(* IEC 61131-3 sources: 2026_Projet_YGO_ExcavatriceDragage/ARCHIVES/Code/PLC_TESTS/CORE, 6 files *)

(* ---- FB_TranslationReportFinalizer.st ---- *)
// ═══════════════════════════════════════════════════════════════
// 🧪 FB_TranslationReportFinalizer — Rapport incrémental Translation
// ───────────────────────────────────────────────────────────────
// 🎯 Responsabilité UNIQUE : enregistrer les verdicts réels et finaliser
//    un rapport borné. Aucun parcours du graphe de transitions.
// ═══════════════════════════════════════════════════════════════

FUNCTION_BLOCK PUBLIC FB_TranslationReportFinalizer
VAR_INPUT
    RunStart        : BOOL;
    RequestedCaseId : INT;
    Busy            : BOOL;
    StepVerdict         : BOOL;
    StepId              : INT;
    StepCaseId          : INT;
    StepPassed          : BOOL;
    StepFailReason      : E_TestFailReason;
    StepFailedCheckIdx  : INT;
    StepDuration        : TIME;
    StepObservedBool    : BOOL;
    StepObservedDint    : DINT;
    StepObservedReal    : REAL;
    Finalize       : BOOL;
    TerminalState  : E_TestTerminalState;
    ErrorCode      : INT;
    ErrorMessage   : STRING(160);
END_VAR
VAR_IN_OUT
    StepTable : ARRAY[1..GVL_PLC_Tests_Const.MaxSteps]     OF ST_TestStepConfig;
    CaseTable : ARRAY[1..GVL_PLC_Tests_Const.MaxTestCases] OF ST_TestCaseConfig;
    Report    : ST_TestSuiteReport;
    Result    : ST_TranslationTestResult;
END_VAR
VAR
    Idx             : INT;
    CaseIdx         : INT;
    CasesTotalLocal : INT;
    CasesPassedLocal: INT;
    CasesFailedLocal: INT;
    FirstFailedCase : INT;
    ReasonText      : STRING(20);
    EntryText       : STRING(80);
END_VAR
// === IMPLEMENTATION ===
IF RunStart THEN
    Report.Name := 'Translation Validation';
    Report.InProgress := TRUE;
    Report.AllPassed := FALSE;
    Report.AnyFailed := FALSE;
    Report.Aborted := FALSE;
    Report.TerminalState := E_TestTerminalState.TEST_TERMINAL_NONE;
    Report.ErrorCode := 0;
    Report.ErrorMessage := '';
    Report.FailedTestCase := 0;
    Report.FailureSummary := '';
    Report.CurrentStepId := 0;
    Report.CurrentCaseId := 0;
    Report.Duration := T#0s;
    Report.RunCounter := Report.RunCounter + 1;
    FOR Idx := 1 TO GVL_PLC_Tests_Const.MaxSteps DO
        Report.Steps[Idx].Executed := FALSE;
        Report.Steps[Idx].Passed := FALSE;
        Report.Steps[Idx].FailReason := E_TestFailReason.FAIL_NONE;
        Report.Steps[Idx].FailedCheckIdx := 0;
        Report.Steps[Idx].FailedInvariantId := 0;
        Report.Steps[Idx].Duration := T#0s;
    END_FOR;
    FOR Idx := 1 TO GVL_PLC_Tests_Const.MaxTestCases DO
        Report.Cases[Idx].Name := CaseTable[Idx].Name;
        Report.Cases[Idx].Executed := FALSE;
        Report.Cases[Idx].Ok := FALSE;
        Report.Cases[Idx].FailedStepId := 0;
        Report.Cases[Idx].FailReason := E_TestFailReason.FAIL_NONE;
        Report.Cases[Idx].Duration := T#0s;
    END_FOR;
    Result.TerminalState := E_TestTerminalState.TEST_TERMINAL_NONE;
    Result.RequestedCaseId := RequestedCaseId;
    Result.ExecutedCaseId := 0;
    Result.AllPassed := FALSE;
    Result.AnyFailed := FALSE;
    Result.FailedCaseId := 0;
    Result.FailedCaseName := '';
    Result.FailReason := E_TestFailReason.FAIL_NONE;
    Result.ErrorCode := 0;
    Result.ErrorMessage := '';
    Result.CasesTotal := 0;
    Result.CasesPassed := 0;
    Result.CasesFailed := 0;
    Result.Duration := T#0s;
    Result.RunCounter := Report.RunCounter;
END_IF;

IF Busy THEN
    Report.Duration := Report.Duration + UDINT_TO_TIME(INT_TO_UDINT(GVL_PLC_Tests_Const.TaskCycleMs));
END_IF;

// 🧾 Agrégation incrémentale : validation séparée avant toute indexation.
IF StepVerdict THEN
    IF StepId < 1 OR StepId > GVL_PLC_Tests_Const.MaxSteps THEN
        Report.ErrorCode := 1050;
        Report.ErrorMessage := 'Verdict StepId hors limites';
        Report.AnyFailed := TRUE;
        RETURN;
    END_IF;
    Report.Steps[StepId].Executed := TRUE;
    Report.Steps[StepId].Passed := StepPassed;
    Report.Steps[StepId].FailReason := StepFailReason;
    Report.Steps[StepId].FailedCheckIdx := StepFailedCheckIdx;
    Report.Steps[StepId].Duration := StepDuration;
    Report.Steps[StepId].ObservedBool := StepObservedBool;
    Report.Steps[StepId].ObservedDint := StepObservedDint;
    Report.Steps[StepId].ObservedReal := StepObservedReal;
    Report.CurrentStepId := StepId;
    Report.CurrentCaseId := StepCaseId;

    IF StepCaseId >= 1 THEN
        IF StepCaseId <= GVL_PLC_Tests_Const.MaxTestCases THEN
        IF NOT Report.Cases[StepCaseId].Executed THEN
            Report.Cases[StepCaseId].Executed := TRUE;
            Report.Cases[StepCaseId].Ok := TRUE;
        END_IF;
        Report.Cases[StepCaseId].Duration := Report.Cases[StepCaseId].Duration + StepDuration;
        IF NOT StepPassed THEN
            Report.Cases[StepCaseId].Ok := FALSE;
            IF Report.Cases[StepCaseId].FailedStepId = 0 THEN
                Report.Cases[StepCaseId].FailedStepId := StepId;
                Report.Cases[StepCaseId].FailReason := StepFailReason;
            END_IF;
        END_IF;
        ELSE
            Report.ErrorCode := 1051;
            Report.ErrorMessage := 'Verdict CaseId hors limites';
            Report.AnyFailed := TRUE;
        END_IF;
    ELSE
        Report.ErrorCode := 1051;
        Report.ErrorMessage := 'Verdict CaseId hors limites';
        Report.AnyFailed := TRUE;
    END_IF;
END_IF;

IF Finalize THEN
    Report.InProgress := FALSE;
    Report.TerminalState := TerminalState;
    Report.ErrorCode := ErrorCode;
    Report.ErrorMessage := ErrorMessage;
    Report.Aborted := (TerminalState = E_TestTerminalState.TEST_TERMINAL_ABORTED);
    CasesTotalLocal := 0;
    CasesPassedLocal := 0;
    CasesFailedLocal := 0;
    FirstFailedCase := 0;
    Report.FailureSummary := '';

    FOR CaseIdx := 1 TO GVL_PLC_Tests_Const.MaxTestCases DO
        IF Report.Cases[CaseIdx].Executed THEN
            CasesTotalLocal := CasesTotalLocal + 1;
            IF Report.Cases[CaseIdx].Ok THEN
                CasesPassedLocal := CasesPassedLocal + 1;
            ELSE
                CasesFailedLocal := CasesFailedLocal + 1;
                IF FirstFailedCase = 0 THEN FirstFailedCase := CaseIdx; END_IF;
                CASE Report.Cases[CaseIdx].FailReason OF
                    E_TestFailReason.FAIL_TIMEOUT: ReasonText := 'FAIL_TIMEOUT';
                    E_TestFailReason.FAIL_CHECK: ReasonText := 'FAIL_CHECK';
                    E_TestFailReason.FAIL_INVARIANT: ReasonText := 'FAIL_INVARIANT';
                    E_TestFailReason.FAIL_WINDOW_EARLY: ReasonText := 'FAIL_WINDOW_EARLY';
                    E_TestFailReason.FAIL_ABORTED: ReasonText := 'FAIL_ABORTED';
                ELSE ReasonText := 'FAIL_NONE';
                END_CASE;
                EntryText := CONCAT(Report.Cases[CaseIdx].Name, ' (step ');
                EntryText := CONCAT(EntryText, INT_TO_STRING(Report.Cases[CaseIdx].FailedStepId));
                EntryText := CONCAT(EntryText, '): ');
                EntryText := CONCAT(EntryText, ReasonText);
                IF Report.FailureSummary = '' THEN
                    Report.FailureSummary := EntryText;
                ELSE
                    Report.FailureSummary := CONCAT(Report.FailureSummary, ' | ');
                    Report.FailureSummary := CONCAT(Report.FailureSummary, EntryText);
                END_IF;
            END_IF;
        END_IF;
    END_FOR;

    Report.AllPassed := (TerminalState = E_TestTerminalState.TEST_TERMINAL_DONE)
                     AND (CasesTotalLocal > 0)
                     AND (CasesFailedLocal = 0);
    Report.AnyFailed := NOT Report.AllPassed;
    Report.FailedTestCase := FirstFailedCase;

    Result.TerminalState := TerminalState;
    Result.RequestedCaseId := RequestedCaseId;
    Result.ExecutedCaseId := Report.CurrentCaseId;
    Result.AllPassed := Report.AllPassed;
    Result.AnyFailed := Report.AnyFailed;
    Result.FailedCaseId := FirstFailedCase;
    IF FirstFailedCase > 0 THEN
        Result.FailedCaseName := Report.Cases[FirstFailedCase].Name;
        Result.FailReason := Report.Cases[FirstFailedCase].FailReason;
    ELSE
        Result.FailedCaseName := '';
        Result.FailReason := E_TestFailReason.FAIL_NONE;
    END_IF;
    Result.ErrorCode := ErrorCode;
    Result.ErrorMessage := ErrorMessage;
    Result.CasesTotal := CasesTotalLocal;
    Result.CasesPassed := CasesPassedLocal;
    Result.CasesFailed := CasesFailedLocal;
    Result.Duration := Report.Duration;
    Result.RunCounter := Report.RunCounter;
END_IF;

(* ---- FB_TranslationStepExecutor.st ---- *)
// ═══════════════════════════════════════════════════════════════
// 🧪 FB_TranslationStepExecutor — Exécution étape/check Translation M3
// ───────────────────────────────────────────────────────────────
// 🎯 Responsabilité UNIQUE : faire progresser UNE suite de tests
//    Translation, étape par étape (Dwell → Checks → Timeout/MinPT →
//    verdict → étape suivante), en respectant le cantonnement à un
//    seul cas (CaseId 1..6) ou à l'enchaînement complet (CaseId=0).
//    N'écrit AUCUNE variable GVL, ne construit AUCUNE table (voir
//    FB_TranslationTestPlan) et n'assemble AUCUN rapport (voir
//    FB_TranslationReportFinalizer, qui consomme StepVerdict/Verdict*).
// 🆕 Tranche verticale NEUVE Translation (2026-07-22) — n'instancie NI
//    FB_TestSequencer NI FB_TestCheck/FB_Timeout (anciennes BRICKS) :
//    logique de check réécrite ici, restreinte aux 3 Kind / 2 Mode
//    réellement utilisés par les 6 TC Translation (voir FB_TranslationTestPlan).
// 🔒 Cantonnement de cas (remplace le FirstStepId manipulé par le
//    manager, audit v1.0 C2) : CaseId est résolu en 1er step via
//    CaseTable UNIQUEMENT ici (jamais exposé par FB_TranslationValidation).
//    Toute étape suivante qui change de CaseId alors qu'un cas est
//    ciblé (CaseId<>0) termine proprement le run (NextStepId:=0).
// ═══════════════════════════════════════════════════════════════

FUNCTION_BLOCK PUBLIC FB_TranslationStepExecutor
VAR_INPUT
    Start   : BOOL; // Front : résout CaseId -> 1er step (CaseTable) et démarre
    Abort   : BOOL; // Niveau : arrêt immédiat propre
    CaseId  : INT;  // 0 = toutes les cases (1..6) ; 1..6 = case ciblée uniquement
END_VAR
VAR_IN_OUT
    StepTable  : ARRAY[1..GVL_PLC_Tests_Const.MaxSteps]      OF ST_TestStepConfig;
    CheckTable : ARRAY[1..GVL_PLC_Tests_Const.MaxChecks]     OF ST_TestCheckConfig;
    CaseTable  : ARRAY[1..GVL_PLC_Tests_Const.MaxTestCases]  OF ST_TestCaseConfig;
    ProbeBool  : ARRAY[1..GVL_PLC_Tests_Const.MaxProbeBool]  OF BOOL;
    ProbeDint  : ARRAY[1..GVL_PLC_Tests_Const.MaxProbeDint]  OF DINT;
    ProbeReal  : ARRAY[1..GVL_PLC_Tests_Const.MaxProbeReal]  OF REAL;
END_VAR
VAR_OUTPUT
    Busy                : BOOL;
    RunDone              : BOOL;  // Fin de run (niveau, tenu jusqu'au prochain Start)
    AnyFailed            : BOOL;
    ConfigError          : BOOL;  // 🛡️ Garde-fou runtime (Plan valide déjà statiquement)
    ConfigErrorStepId    : INT;
    CurrentStepId        : INT;
    CurrentCaseId        : INT;
    ActiveStimulusId     : INT;   // 0 GARANTI sur tout chemin terminal (Done/Abort/ConfigError)
    StepElapsed          : TIME;
    TerminalState        : E_TestTerminalState;
    // 🧾 Verdict d'étape — pulse 1 scan, consommé par FB_TranslationReportFinalizer
    StepVerdict          : BOOL;
    VerdictStepId        : INT;
    VerdictCaseId        : INT;
    VerdictPassed         : BOOL;
    VerdictFailReason     : E_TestFailReason;
    VerdictFailedCheckIdx : INT;
    VerdictDuration       : TIME;
    VerdictObservedBool   : BOOL;
    VerdictObservedDint   : DINT;
    VerdictObservedReal   : REAL;
END_VAR
VAR
    StartTrig       : R_TRIG;
    StepStarted     : BOOL;
    DwellTimer      : TON;
    StepTimer       : TON;
    StableTimers    : ARRAY[1..GVL_PLC_Tests_Const.MaxChecksPerStep] OF TON;
    CheckPassed     : ARRAY[1..GVL_PLC_Tests_Const.MaxChecksPerStep] OF BOOL;
    CheckFailed     : ARRAY[1..GVL_PLC_Tests_Const.MaxChecksPerStep] OF BOOL;
    InstantEvaluated: ARRAY[1..GVL_PLC_Tests_Const.MaxChecksPerStep] OF BOOL;
    ObsBoolArr      : ARRAY[1..GVL_PLC_Tests_Const.MaxChecksPerStep] OF BOOL;
    ObsDintArr      : ARRAY[1..GVL_PLC_Tests_Const.MaxChecksPerStep] OF DINT;
    ObsRealArr      : ARRAY[1..GVL_PLC_Tests_Const.MaxChecksPerStep] OF REAL;

    Jdx, Kdx        : INT;
    ProbeIdx        : INT;
    Cond            : BOOL;
    AllChecksLatched: BOOL;
    AnyCheckFailedLocal : BOOL;
    FailedCheckIdxLocal : INT;
    FailedCheckSlotLocal : INT; // Slot RÉEL (Jdx, 1..MaxChecksPerStep) du check fautif

    // Verdict de l'étape (émis au plus une fois par scan)
    VerdictReached      : BOOL;
    VerdictPassedLocal   : BOOL;
    VerdictReasonLocal   : E_TestFailReason;
    VerdictCheckIdxLocal : INT;
    VerdictObsBoolLocal  : BOOL;
    VerdictObsDintLocal  : DINT;
    VerdictObsRealLocal  : REAL;

    NextCandidate    : INT;
    TransitionCount  : INT; // Garde anti-cycle runtime, bornée par MaxSteps
END_VAR
// === IMPLEMENTATION ===
StartTrig(CLK := Start);
StepVerdict := FALSE;

// 1. 🛑 Abort — niveau, priorité absolue
IF Abort THEN
    IF Busy THEN
        StepVerdict := TRUE;
        VerdictStepId := CurrentStepId;
        VerdictCaseId := CurrentCaseId;
        VerdictPassed := FALSE;
        VerdictFailReason := E_TestFailReason.FAIL_ABORTED;
        VerdictFailedCheckIdx := 0;
        VerdictDuration := StepElapsed;
        VerdictObservedBool := FALSE;
        VerdictObservedDint := 0;
        VerdictObservedReal := 0.0;
        AnyFailed := TRUE;
        TerminalState := E_TestTerminalState.TEST_TERMINAL_ABORTED;
    END_IF;
    Busy := FALSE;
    RunDone := TRUE;
    ActiveStimulusId := 0;
    CurrentStepId := 0;
    StepStarted := FALSE;
    RETURN;
END_IF;

// 2. 🟢 Démarrage — résolution CaseId -> 1er step, JAMAIS de FirstStepId externe
IF StartTrig.Q THEN
    ConfigError := FALSE;
    ConfigErrorStepId := 0;
    TerminalState := E_TestTerminalState.TEST_TERMINAL_NONE;

    IF CaseId < 0 OR CaseId > 6 THEN
        ConfigError := TRUE;
        ConfigErrorStepId := CaseId;
        Busy := FALSE;
        RunDone := TRUE;
        AnyFailed := TRUE;
        ActiveStimulusId := 0;
        CurrentStepId := 0;
        TerminalState := E_TestTerminalState.TEST_TERMINAL_CONFIG_ERROR;
        RETURN;
    END_IF;

    IF CaseId = 0 THEN
        CurrentStepId := CaseTable[1].FirstStep;
    ELSE
        CurrentStepId := CaseTable[CaseId].FirstStep;
    END_IF;

    IF CurrentStepId < 1 OR CurrentStepId > GVL_PLC_Tests_Const.MaxSteps THEN
        ConfigError := TRUE;
        ConfigErrorStepId := CurrentStepId;
        Busy := FALSE;
        RunDone := TRUE;
        AnyFailed := TRUE;
        ActiveStimulusId := 0;
        CurrentStepId := 0;
        TerminalState := E_TestTerminalState.TEST_TERMINAL_CONFIG_ERROR;
        RETURN;
    END_IF;

    Busy := TRUE;
    RunDone := FALSE;
    AnyFailed := FALSE;
    StepStarted := FALSE;
    TransitionCount := 0;
END_IF;

IF NOT Busy THEN
    RETURN;
END_IF;

// 3. 🛡️ Garde-fou runtime (défense en profondeur — Plan valide déjà statiquement)
IF CurrentStepId < 1 OR CurrentStepId > GVL_PLC_Tests_Const.MaxSteps THEN
    Busy := FALSE;
    RunDone := TRUE;
    AnyFailed := TRUE;
    ActiveStimulusId := 0;
    ConfigError := TRUE;
    ConfigErrorStepId := CurrentStepId;
    TerminalState := E_TestTerminalState.TEST_TERMINAL_CONFIG_ERROR;
    RETURN;
END_IF;

CurrentCaseId := StepTable[CurrentStepId].CaseId;
ActiveStimulusId := StepTable[CurrentStepId].StimulusId;

IF NOT StepStarted THEN
    StepStarted := TRUE;
    StepElapsed := T#0s;
    DwellTimer(IN := FALSE);
    StepTimer(IN := FALSE);
    FOR Jdx := 1 TO GVL_PLC_Tests_Const.MaxChecksPerStep DO
        CheckPassed[Jdx] := FALSE;
        CheckFailed[Jdx] := FALSE;
        InstantEvaluated[Jdx] := FALSE;
        StableTimers[Jdx](IN := FALSE);
    END_FOR;
END_IF;

StepElapsed := StepElapsed + UDINT_TO_TIME(INT_TO_UDINT(GVL_PLC_Tests_Const.TaskCycleMs));

// 4. 🕐 Dwell (tempo fixe avant évaluation — T#0s = aucune, cas actuel Translation)
DwellTimer(IN := TRUE, PT := StepTable[CurrentStepId].DwellPT);
IF NOT DwellTimer.Q THEN
    RETURN;
END_IF;

// 5. ✅ Évaluation des checks — verrouillage "latch and hold" par check
//    (un check WAIT_UNTIL passé le reste jusqu'à la fin de l'étape, même si
//    la sonde redevient momentanément fausse — sémantique identique à
//    l'ancien FB_TestCheck, réécrite ici sans l'instancier)
FOR Jdx := 1 TO GVL_PLC_Tests_Const.MaxChecksPerStep DO
    Kdx := StepTable[CurrentStepId].CheckIdx[Jdx];
    // 🔒 CODESYS n'assure pas le court-circuit : valider AVANT tout accès.
    IF Kdx < 0 OR Kdx > GVL_PLC_Tests_Const.MaxChecks THEN
        Busy := FALSE;
        RunDone := TRUE;
        AnyFailed := TRUE;
        ActiveStimulusId := 0;
        ConfigError := TRUE;
        ConfigErrorStepId := CurrentStepId;
        TerminalState := E_TestTerminalState.TEST_TERMINAL_CONFIG_ERROR;
        RETURN;
    END_IF;
    IF Kdx > 0 THEN
        Cond := FALSE;
        ProbeIdx := CheckTable[Kdx].ProbeIdx;
        CASE CheckTable[Kdx].Kind OF
            E_TestCheckKind.BOOL_EQUAL:
                IF ProbeIdx >= 1 THEN
                    IF ProbeIdx <= GVL_PLC_Tests_Const.MaxProbeBool THEN
                        ObsBoolArr[Jdx] := ProbeBool[ProbeIdx];
                        Cond := (ObsBoolArr[Jdx] = CheckTable[Kdx].ExpectedBool);
                    END_IF;
                END_IF;
            E_TestCheckKind.WORD_MASK_NONE:
                IF ProbeIdx >= 1 THEN
                    IF ProbeIdx <= GVL_PLC_Tests_Const.MaxProbeDint THEN
                        ObsDintArr[Jdx] := ProbeDint[ProbeIdx];
                        Cond := ((DINT_TO_WORD(ObsDintArr[Jdx]) AND CheckTable[Kdx].Mask) = 0);
                    END_IF;
                END_IF;
            E_TestCheckKind.REAL_IN_RANGE:
                IF ProbeIdx >= 1 THEN
                    IF ProbeIdx <= GVL_PLC_Tests_Const.MaxProbeReal THEN
                        ObsRealArr[Jdx] := ProbeReal[ProbeIdx];
                        Cond := (ObsRealArr[Jdx] >= CheckTable[Kdx].RealMin AND ObsRealArr[Jdx] <= CheckTable[Kdx].RealMax);
                    END_IF;
                END_IF;
            // Kind hors périmètre (voir FB_TranslationTestPlan) -> Cond reste FALSE
        END_CASE;

        IF NOT CheckPassed[Jdx] AND NOT CheckFailed[Jdx] THEN
            CASE CheckTable[Kdx].Mode OF
                E_TestCheckMode.CHECK_INSTANT:
                    IF NOT InstantEvaluated[Jdx] THEN
                        InstantEvaluated[Jdx] := TRUE;
                        IF Cond THEN
                            CheckPassed[Jdx] := TRUE;
                        ELSE
                            CheckFailed[Jdx] := TRUE;
                        END_IF;
                    END_IF;
                E_TestCheckMode.CHECK_WAIT_UNTIL:
                    StableTimers[Jdx](IN := Cond, PT := CheckTable[Kdx].StablePT);
                    IF StableTimers[Jdx].Q THEN
                        CheckPassed[Jdx] := TRUE;
                    END_IF;
            END_CASE;
        END_IF;
    END_IF;
END_FOR;

// 6. 🧾 Agrégat des checks de l'étape
AllChecksLatched := TRUE;
AnyCheckFailedLocal := FALSE;
FailedCheckIdxLocal := 0;
FailedCheckSlotLocal := 0;
FOR Jdx := 1 TO GVL_PLC_Tests_Const.MaxChecksPerStep DO
    Kdx := StepTable[CurrentStepId].CheckIdx[Jdx];
    IF Kdx > 0 THEN
        IF CheckFailed[Jdx] AND NOT AnyCheckFailedLocal THEN
            AnyCheckFailedLocal := TRUE;
            FailedCheckIdxLocal := Kdx;
            FailedCheckSlotLocal := Jdx; // 🔧 REX : slot RÉEL du check fautif (pas un index figé)
        ELSIF NOT CheckPassed[Jdx] THEN
            AllChecksLatched := FALSE;
        END_IF;
    END_IF;
END_FOR;

// 7. 📸 Verdict
VerdictReached := FALSE;
IF AnyCheckFailedLocal THEN
    VerdictReached := TRUE;
    VerdictPassedLocal := FALSE;
    VerdictReasonLocal := E_TestFailReason.FAIL_CHECK;
    VerdictCheckIdxLocal := FailedCheckIdxLocal;
    // 🔒 Défense en profondeur avant indexation du snapshot fautif.
    IF FailedCheckSlotLocal >= 1 THEN
        IF FailedCheckSlotLocal <= GVL_PLC_Tests_Const.MaxChecksPerStep THEN
            VerdictObsBoolLocal := ObsBoolArr[FailedCheckSlotLocal];
            VerdictObsDintLocal := ObsDintArr[FailedCheckSlotLocal];
            VerdictObsRealLocal := ObsRealArr[FailedCheckSlotLocal];
        ELSE
            VerdictObsBoolLocal := FALSE;
            VerdictObsDintLocal := 0;
            VerdictObsRealLocal := 0.0;
        END_IF;
    ELSE
        VerdictObsBoolLocal := FALSE;
        VerdictObsDintLocal := 0;
        VerdictObsRealLocal := 0.0;
    END_IF;
ELSE
    StepTimer(IN := TRUE, PT := StepTable[CurrentStepId].TimeoutPT);
    IF AllChecksLatched THEN
        VerdictReached := TRUE;
        IF StepElapsed < StepTable[CurrentStepId].MinPT THEN
            VerdictPassedLocal := FALSE;
            VerdictReasonLocal := E_TestFailReason.FAIL_WINDOW_EARLY;
            VerdictCheckIdxLocal := 0;
        ELSE
            VerdictPassedLocal := TRUE;
            VerdictReasonLocal := E_TestFailReason.FAIL_NONE;
            VerdictCheckIdxLocal := 0;
        END_IF;
        VerdictObsBoolLocal := ObsBoolArr[1];
        VerdictObsDintLocal := ObsDintArr[1];
        VerdictObsRealLocal := ObsRealArr[1];
    ELSIF StepTimer.Q THEN
        VerdictReached := TRUE;
        VerdictPassedLocal := FALSE;
        VerdictReasonLocal := E_TestFailReason.FAIL_TIMEOUT;
        VerdictCheckIdxLocal := 0;
        VerdictObsBoolLocal := FALSE;
        VerdictObsDintLocal := 0;
        VerdictObsRealLocal := 0.0;
    END_IF;
END_IF;

IF NOT VerdictReached THEN
    RETURN; // ⏳ Toujours en attente, rien à publier ce scan
END_IF;

// 8. ➡️ Résolution de l'étape suivante — cantonnement de cas ICI (audit v1.0 C2)
IF VerdictPassedLocal THEN
    NextCandidate := StepTable[CurrentStepId].NextOnPass;
ELSIF StepTable[CurrentStepId].FailAction = E_TestFailAction.FAIL_ABORT_SUITE THEN
    NextCandidate := 0;
ELSE
    NextCandidate := StepTable[CurrentStepId].NextOnFail;
END_IF;

// 🔒 Aucun accès StepTable[0] : CODESYS peut évaluer tous les opérandes de AND.
IF NextCandidate <> 0 THEN
    IF NextCandidate < 1 OR NextCandidate > GVL_PLC_Tests_Const.MaxSteps THEN
        Busy := FALSE;
        RunDone := TRUE;
        AnyFailed := TRUE;
        ActiveStimulusId := 0;
        ConfigError := TRUE;
        ConfigErrorStepId := NextCandidate;
        TerminalState := E_TestTerminalState.TEST_TERMINAL_CONFIG_ERROR;
        RETURN;
    END_IF;
    // Un cas ciblé ne déborde jamais sur le cas suivant.
    IF CaseId <> 0 THEN
        IF StepTable[NextCandidate].CaseId <> CaseId THEN
            NextCandidate := 0;
        END_IF;
    END_IF;
END_IF;

// 9. 🧾 Publication du verdict pour FB_TranslationReportFinalizer
StepVerdict := TRUE;
VerdictStepId := CurrentStepId;
VerdictCaseId := CurrentCaseId;
VerdictPassed := VerdictPassedLocal;
VerdictFailReason := VerdictReasonLocal;
VerdictFailedCheckIdx := VerdictCheckIdxLocal;
VerdictDuration := StepElapsed;
VerdictObservedBool := VerdictObsBoolLocal;
VerdictObservedDint := VerdictObsDintLocal;
VerdictObservedReal := VerdictObsRealLocal;

IF NOT VerdictPassedLocal THEN
    AnyFailed := TRUE;
END_IF;

// 10. 🔁 Transition bornée (garde runtime contre tout cycle résiduel)
TransitionCount := TransitionCount + 1;
IF TransitionCount > GVL_PLC_Tests_Const.MaxSteps THEN
    Busy := FALSE;
    RunDone := TRUE;
    AnyFailed := TRUE;
    ActiveStimulusId := 0;
    ConfigError := TRUE;
    ConfigErrorStepId := CurrentStepId;
    TerminalState := E_TestTerminalState.TEST_TERMINAL_CONFIG_ERROR;
    RETURN;
END_IF;
CurrentStepId := NextCandidate;
StepStarted := FALSE;
IF NextCandidate = 0 THEN
    Busy := FALSE;
    RunDone := TRUE;
    ActiveStimulusId := 0; // 🛡️ Garantie structurelle — double garantie avec FB_TranslationTestCleanup
    IF AnyFailed THEN
        TerminalState := E_TestTerminalState.TEST_TERMINAL_FAILED;
    ELSE
        TerminalState := E_TestTerminalState.TEST_TERMINAL_DONE;
    END_IF;
END_IF;

(* ---- FB_TranslationTestCleanup.st ---- *)
// ═══════════════════════════════════════════════════════════════
// 🧪 FB_TranslationTestCleanup — Neutralité Translation M3
// ───────────────────────────────────────────────────────────────
// 🎯 Responsabilité UNIQUE : porter le vecteur d'état NEUTRE complet
//    (tous les overrides M3 relâchés, instance isolée FB_Translation
//    au repos). Source de vérité UNIQUE de "neutre" — appelée depuis
//    le fichier suite (SUITE_TRANSLATION/FB_TranslationValidation.st)
//    à la fois dans le CASE stimulus (StimulusId=0) ET, en garantie
//    structurelle indépendante, sur tout chemin où la suite n'est pas
//    Busy (ceinture + bretelles, AF_Partie-14 §7.3.2).
// 🚫 Ne force JAMAIS une sortie de commande calculée — uniquement les
//    surcharges capteurs amont (GVL_PLC_Tests.OverrideM3*) et les
//    entrées de l'instance de test isolée.
// ═══════════════════════════════════════════════════════════════

FUNCTION_BLOCK PUBLIC FB_TranslationTestCleanup
VAR_INPUT
    Apply : BOOL; // TRUE = force la neutralité maintenant
END_VAR
VAR_OUTPUT
    OverrideAtTremie          : BOOL;
    OverrideBrakeStuckOpen    : BOOL;
    OverridePhantomFreq       : BOOL;
    OverrideSensorsWordActive : BOOL;
    UnderTestDirection        : INT;
    UnderTestStartStop        : BOOL;
    UnderTestSlowdownSensor   : BOOL;
    NeutralConfirmed          : BOOL; // TRUE dès que la neutralité a été appliquée ce scan
END_VAR
// === IMPLEMENTATION ===
IF Apply THEN
    OverrideAtTremie := FALSE;
    OverrideBrakeStuckOpen := FALSE;
    OverridePhantomFreq := FALSE;
    OverrideSensorsWordActive := FALSE;
    UnderTestDirection := 0;
    UnderTestStartStop := FALSE;
    UnderTestSlowdownSensor := FALSE;
    NeutralConfirmed := TRUE;
ELSE
    NeutralConfirmed := FALSE;
END_IF;

(* ---- FB_TranslationTestFixture.st ---- *)
// ═══════════════════════════════════════════════════════════════
// 🧪 FB_TranslationTestFixture — Précondition Translation M3
// ───────────────────────────────────────────────────────────────
// 🎯 Responsabilité UNIQUE : décider si un Start est recevable
//    (Niveaux 1/2 de la défense en profondeur, AF_Partie-14 §7.3.3) :
//    simulation active + aucune E/S M3 recâblée réelle. Ne fait AUCUNE
//    attente d'état sain (ça reste la responsabilité de l'étape SETUP
//    de chaque cas, via FB_TranslationStepExecutor — §7.3.5).
// 🔒 Un refus ici est TOUJOURS explicite (PRECONDITION_FAILED),
//    jamais un silence (audit v1.0 C3).
// ═══════════════════════════════════════════════════════════════

FUNCTION_BLOCK PUBLIC FB_TranslationTestFixture
VAR_INPUT
    CheckRequested        : BOOL; // Front : nouvelle vérification demandée (sur Start suite)
    SimulationModeActive  : BOOL;
    SimGateOk             : BOOL; // Niveau 2 : aucune E/S M3 (*IsReal) incompatible
END_VAR
VAR_OUTPUT
    FixturePassed  : BOOL;
    FixtureFailed  : BOOL;
    FailReason     : STRING(120);
END_VAR
VAR
    CheckTrig : R_TRIG;
END_VAR
// === IMPLEMENTATION ===
CheckTrig(CLK := CheckRequested);

IF CheckTrig.Q THEN
    IF NOT SimulationModeActive THEN
        FixturePassed := FALSE;
        FixtureFailed := TRUE;
        FailReason := 'Simulation non active (GVL_Simulation.SimulationModeActive=FALSE)';
    ELSIF NOT SimGateOk THEN
        FixturePassed := FALSE;
        FixtureFailed := TRUE;
        FailReason := 'E/S M3 recablees reelles (*IsReal) incompatibles avec le banc de test';
    ELSE
        FixturePassed := TRUE;
        FixtureFailed := FALSE;
        FailReason := '';
    END_IF;
END_IF;

(* ---- FB_TranslationTestPlan.st ---- *)
// ═══════════════════════════════════════════════════════════════
// 🧪 FB_TranslationTestPlan — Plan de validation Translation M3
// ───────────────────────────────────────────────────────────────
// 🎯 Responsabilité UNIQUE : construire (une seule fois) et auto-valider
//    les tables déclaratives (StepTable/CheckTable/CaseTable) de la
//    suite Translation, puis exposer un refus explicite ConfigError si
//    la table est incohérente. Ne pilote AUCUNE exécution (voir
//    FB_TranslationStepExecutor) et n'écrit AUCUNE variable GVL.
// 🆕 Tranche verticale NEUVE Translation (2026-07-22) — moteur dédié,
//    n'instancie NI FB_TestSequencer NI les anciennes BRICKS
//    (FB_TestCheck/FB_Timeout...). Voir DOC/AUDITS/TEST_FRAMEWORK_AUDIT_v1.0.md.
// 📌 Périmètre volontairement restreint (audit §"strictement nécessaires") :
//    seuls les Kind/Mode réellement utilisés par les 6 TC Translation
//    sont acceptés — BOOL_EQUAL/WORD_MASK_NONE/REAL_IN_RANGE,
//    CHECK_INSTANT/CHECK_WAIT_UNTIL. Tout autre Kind/Mode -> ConfigError.
// 🔑 Index des sondes (Sig*) : PLUS possédés ici. Le fichier suite
//    (SUITE_TRANSLATION/FB_TranslationValidation.st) les déclare comme
//    SES PROPRES VAR CONSTANT et les transmet en VAR_INPUT à chaque appel
//    -- aucun accès croisé "instPlan.SigXxx" depuis l'extérieur. Le Plan
//    ne fait que les recopier dans CheckTable[].ProbeIdx à la construction.
// ═══════════════════════════════════════════════════════════════

FUNCTION_BLOCK PUBLIC FB_TranslationTestPlan
VAR_INPUT
    // 🏷️ Index des sondes — fournis par l'appelant (source de vérité :
    //    VAR CONSTANT de FB_TranslationValidation), jamais lus en retour.
    SigHealthyIdle          : INT;
    SigLimitSwitchError     : INT;
    SigPowerCutOff          : INT;
    SigErrorIdT1NoParasite  : INT;
    SigMecaBError            : INT;
    SigErrorIdT2NoParasite  : INT;
    SigMecaAError            : INT;
    SigErrorIdT3NoParasite  : INT;
    SigDecoderIncoherent     : INT;
    SigLimitFwd              : INT;
    SigLimitRev              : INT;
    SigSensorIncoherentErr  : INT;
    SigErrorIdT5NoParasite  : INT; // DINT
    SigSlowdownFreqHz        : INT; // REAL
END_VAR
VAR_OUTPUT
    Ready               : BOOL;   // Tables construites + validées
    ConfigError          : BOOL;  // 🔒 Table invalide -> aucun Start ne doit être honoré
    ConfigErrorStepId    : INT;
    ConfigErrorCheckIdx  : INT;
    ConfigErrorMessage   : STRING(160);
END_VAR
VAR_IN_OUT
    StepTable  : ARRAY[1..GVL_PLC_Tests_Const.MaxSteps]      OF ST_TestStepConfig;
    CheckTable : ARRAY[1..GVL_PLC_Tests_Const.MaxChecks]     OF ST_TestCheckConfig;
    CaseTable  : ARRAY[1..GVL_PLC_Tests_Const.MaxTestCases]  OF ST_TestCaseConfig;
END_VAR
VAR
    // 🪜 Index des étapes (usage interne uniquement — assemblage des tables)
    StepTc01Setup     : INT := 10;
    StepTc01Trigger   : INT := 11;
    StepTc01Teardown  : INT := 19;

    StepTc02Setup     : INT := 20;
    StepTc02Trigger   : INT := 21;
    StepTc02Teardown  : INT := 29;

    StepTc03Setup     : INT := 30;
    StepTc03Trigger   : INT := 31;
    StepTc03Teardown  : INT := 39;

    StepTc04Setup            : INT := 40;
    StepTc04Word1Tremie      : INT := 41;
    StepTc04Word2            : INT := 42;
    StepTc04Word3            : INT := 43;
    StepTc04Word4            : INT := 44;
    StepTc04Word5             : INT := 45;
    StepTc04Word6Maintenance : INT := 46;
    StepTc04Teardown          : INT := 49;

    StepTc05Setup     : INT := 50;
    StepTc05Trigger   : INT := 51;
    StepTc05Teardown  : INT := 59;

    StepTc06Setup      : INT := 60;
    StepTc06FullSpeed  : INT := 61;
    StepTc06Slowdown   : INT := 62;
    StepTc06Teardown   : INT := 63;

    Built  : BOOL;
    Idx    : INT;
    Jdx    : INT;
    Kdx       : INT;
    WalkIdx   : INT;
    WalkStep  : INT;
    HasCheck  : BOOL;
END_VAR
// === IMPLEMENTATION ===

// 1. 📋 CONSTRUCTION (une seule fois, données pures)
IF NOT Built THEN

    // --- Cas de tests ---
    CaseTable[1].Name := 'TC-T1 Fin de course extreme';
    CaseTable[1].FirstStep := StepTc01Setup;
    CaseTable[2].Name := 'TC-T2 Meca B incoherence arret';
    CaseTable[2].FirstStep := StepTc02Setup;
    CaseTable[3].Name := 'TC-T3 Meca A mvt non commande';
    CaseTable[3].FirstStep := StepTc03Setup;
    CaseTable[4].Name := 'TC-T4 Mots valides + limites';
    CaseTable[4].FirstStep := StepTc04Setup;
    CaseTable[5].Name := 'TC-T5 Incoherence mot capteurs';
    CaseTable[5].FirstStep := StepTc05Setup;
    CaseTable[6].Name := 'TC-T6 Ralentissement PV';
    CaseTable[6].FirstStep := StepTc06Setup;

    // --- Checks ---
    CheckTable[1].Kind := E_TestCheckKind.BOOL_EQUAL;
    CheckTable[1].Mode := E_TestCheckMode.CHECK_WAIT_UNTIL;
    CheckTable[1].ProbeIdx := SigHealthyIdle;
    CheckTable[1].ExpectedBool := TRUE;

    CheckTable[2].Kind := E_TestCheckKind.BOOL_EQUAL;
    CheckTable[2].Mode := E_TestCheckMode.CHECK_WAIT_UNTIL;
    CheckTable[2].ProbeIdx := SigLimitSwitchError;
    CheckTable[2].ExpectedBool := TRUE;

    CheckTable[3].Kind := E_TestCheckKind.BOOL_EQUAL;
    CheckTable[3].Mode := E_TestCheckMode.CHECK_WAIT_UNTIL;
    CheckTable[3].ProbeIdx := SigPowerCutOff;
    CheckTable[3].ExpectedBool := TRUE;

    CheckTable[4].Kind := E_TestCheckKind.WORD_MASK_NONE;
    CheckTable[4].Mode := E_TestCheckMode.CHECK_WAIT_UNTIL;
    CheckTable[4].ProbeIdx := SigErrorIdT1NoParasite;
    CheckTable[4].Mask := NOT 16#0040;

    CheckTable[5].Kind := E_TestCheckKind.BOOL_EQUAL;
    CheckTable[5].Mode := E_TestCheckMode.CHECK_WAIT_UNTIL;
    CheckTable[5].ProbeIdx := SigMecaBError;
    CheckTable[5].ExpectedBool := TRUE;

    CheckTable[6].Kind := E_TestCheckKind.WORD_MASK_NONE;
    CheckTable[6].Mode := E_TestCheckMode.CHECK_WAIT_UNTIL;
    CheckTable[6].ProbeIdx := SigErrorIdT2NoParasite;
    CheckTable[6].Mask := NOT 16#0010;

    CheckTable[7].Kind := E_TestCheckKind.BOOL_EQUAL;
    CheckTable[7].Mode := E_TestCheckMode.CHECK_WAIT_UNTIL;
    CheckTable[7].ProbeIdx := SigMecaAError;
    CheckTable[7].ExpectedBool := TRUE;

    CheckTable[8].Kind := E_TestCheckKind.WORD_MASK_NONE;
    CheckTable[8].Mode := E_TestCheckMode.CHECK_WAIT_UNTIL;
    CheckTable[8].ProbeIdx := SigErrorIdT3NoParasite;
    CheckTable[8].Mask := NOT 16#0020;

    CheckTable[9].Kind := E_TestCheckKind.BOOL_EQUAL;
    CheckTable[9].Mode := E_TestCheckMode.CHECK_WAIT_UNTIL;
    CheckTable[9].ProbeIdx := SigDecoderIncoherent;
    CheckTable[9].ExpectedBool := FALSE;

    CheckTable[10].Kind := E_TestCheckKind.BOOL_EQUAL;
    CheckTable[10].Mode := E_TestCheckMode.CHECK_WAIT_UNTIL;
    CheckTable[10].ProbeIdx := SigLimitFwd;
    CheckTable[10].ExpectedBool := TRUE;

    CheckTable[11].Kind := E_TestCheckKind.BOOL_EQUAL;
    CheckTable[11].Mode := E_TestCheckMode.CHECK_WAIT_UNTIL;
    CheckTable[11].ProbeIdx := SigLimitRev;
    CheckTable[11].ExpectedBool := FALSE;

    CheckTable[12].Kind := E_TestCheckKind.BOOL_EQUAL;
    CheckTable[12].Mode := E_TestCheckMode.CHECK_WAIT_UNTIL;
    CheckTable[12].ProbeIdx := SigLimitRev;
    CheckTable[12].ExpectedBool := TRUE;

    CheckTable[13].Kind := E_TestCheckKind.BOOL_EQUAL;
    CheckTable[13].Mode := E_TestCheckMode.CHECK_WAIT_UNTIL;
    CheckTable[13].ProbeIdx := SigLimitFwd;
    CheckTable[13].ExpectedBool := FALSE;

    CheckTable[14].Kind := E_TestCheckKind.BOOL_EQUAL;
    CheckTable[14].Mode := E_TestCheckMode.CHECK_WAIT_UNTIL;
    CheckTable[14].ProbeIdx := SigLimitFwd;
    CheckTable[14].ExpectedBool := FALSE;

    CheckTable[15].Kind := E_TestCheckKind.BOOL_EQUAL;
    CheckTable[15].Mode := E_TestCheckMode.CHECK_WAIT_UNTIL;
    CheckTable[15].ProbeIdx := SigLimitRev;
    CheckTable[15].ExpectedBool := FALSE;

    CheckTable[16].Kind := E_TestCheckKind.BOOL_EQUAL;
    CheckTable[16].Mode := E_TestCheckMode.CHECK_WAIT_UNTIL;
    CheckTable[16].ProbeIdx := SigDecoderIncoherent;
    CheckTable[16].ExpectedBool := TRUE;

    CheckTable[17].Kind := E_TestCheckKind.BOOL_EQUAL;
    CheckTable[17].Mode := E_TestCheckMode.CHECK_WAIT_UNTIL;
    CheckTable[17].ProbeIdx := SigSensorIncoherentErr;
    CheckTable[17].ExpectedBool := TRUE;

    CheckTable[18].Kind := E_TestCheckKind.WORD_MASK_NONE;
    CheckTable[18].Mode := E_TestCheckMode.CHECK_WAIT_UNTIL;
    CheckTable[18].ProbeIdx := SigErrorIdT5NoParasite;
    CheckTable[18].Mask := NOT 16#0080;

    CheckTable[19].Kind := E_TestCheckKind.REAL_IN_RANGE;
    CheckTable[19].Mode := E_TestCheckMode.CHECK_WAIT_UNTIL;
    CheckTable[19].ProbeIdx := SigSlowdownFreqHz;
    CheckTable[19].RealMin := 30.0;
    CheckTable[19].RealMax := 60.0;

    CheckTable[20].Kind := E_TestCheckKind.REAL_IN_RANGE;
    CheckTable[20].Mode := E_TestCheckMode.CHECK_WAIT_UNTIL;
    CheckTable[20].ProbeIdx := SigSlowdownFreqHz;
    CheckTable[20].RealMin := 8.0;
    CheckTable[20].RealMax := 14.0;

    // --- TC-T1 ---
    StepTable[StepTc01Setup].Name := 'TCT1 Setup saine';
    StepTable[StepTc01Setup].CaseId := 1;
    StepTable[StepTc01Setup].StimulusId := 1;
    StepTable[StepTc01Setup].CheckIdx[1] := 1;
    StepTable[StepTc01Setup].TimeoutPT := T#12s;
    StepTable[StepTc01Setup].NextOnPass := StepTc01Trigger;
    StepTable[StepTc01Setup].NextOnFail := StepTc01Teardown;
    StepTable[StepTc01Setup].FailAction := E_TestFailAction.FAIL_CONTINUE;

    StepTable[StepTc01Trigger].Name := 'TCT1 Fdc Tremie force';
    StepTable[StepTc01Trigger].CaseId := 1;
    StepTable[StepTc01Trigger].StimulusId := 2;
    StepTable[StepTc01Trigger].CheckIdx[1] := 2;
    StepTable[StepTc01Trigger].CheckIdx[2] := 3;
    StepTable[StepTc01Trigger].CheckIdx[3] := 4;
    StepTable[StepTc01Trigger].TimeoutPT := T#5s;
    StepTable[StepTc01Trigger].NextOnPass := StepTc01Teardown;
    StepTable[StepTc01Trigger].NextOnFail := StepTc01Teardown;
    StepTable[StepTc01Trigger].FailAction := E_TestFailAction.FAIL_CONTINUE;

    StepTable[StepTc01Teardown].Name := 'TCT1 Teardown';
    StepTable[StepTc01Teardown].CaseId := 1;
    StepTable[StepTc01Teardown].StimulusId := 1;
    StepTable[StepTc01Teardown].CheckIdx[1] := 1;
    StepTable[StepTc01Teardown].TimeoutPT := T#12s;
    StepTable[StepTc01Teardown].NextOnPass := StepTc02Setup;
    StepTable[StepTc01Teardown].NextOnFail := StepTc02Setup;
    StepTable[StepTc01Teardown].FailAction := E_TestFailAction.FAIL_CONTINUE;

    // --- TC-T2 ---
    StepTable[StepTc02Setup].Name := 'TCT2 Setup saine';
    StepTable[StepTc02Setup].CaseId := 2;
    StepTable[StepTc02Setup].StimulusId := 1;
    StepTable[StepTc02Setup].CheckIdx[1] := 1;
    StepTable[StepTc02Setup].TimeoutPT := T#12s;
    StepTable[StepTc02Setup].NextOnPass := StepTc02Trigger;
    StepTable[StepTc02Setup].NextOnFail := StepTc02Teardown;
    StepTable[StepTc02Setup].FailAction := E_TestFailAction.FAIL_CONTINUE;

    StepTable[StepTc02Trigger].Name := 'TCT2 Frein bloque ouvert';
    StepTable[StepTc02Trigger].CaseId := 2;
    StepTable[StepTc02Trigger].StimulusId := 3;
    StepTable[StepTc02Trigger].CheckIdx[1] := 5;
    StepTable[StepTc02Trigger].CheckIdx[2] := 3;
    StepTable[StepTc02Trigger].CheckIdx[3] := 6;
    StepTable[StepTc02Trigger].TimeoutPT := T#6s;
    StepTable[StepTc02Trigger].NextOnPass := StepTc02Teardown;
    StepTable[StepTc02Trigger].NextOnFail := StepTc02Teardown;
    StepTable[StepTc02Trigger].FailAction := E_TestFailAction.FAIL_CONTINUE;

    StepTable[StepTc02Teardown].Name := 'TCT2 Teardown';
    StepTable[StepTc02Teardown].CaseId := 2;
    StepTable[StepTc02Teardown].StimulusId := 1;
    StepTable[StepTc02Teardown].CheckIdx[1] := 1;
    StepTable[StepTc02Teardown].TimeoutPT := T#12s;
    StepTable[StepTc02Teardown].NextOnPass := StepTc03Setup;
    StepTable[StepTc02Teardown].NextOnFail := StepTc03Setup;
    StepTable[StepTc02Teardown].FailAction := E_TestFailAction.FAIL_CONTINUE;

    // --- TC-T3 ---
    StepTable[StepTc03Setup].Name := 'TCT3 Setup saine';
    StepTable[StepTc03Setup].CaseId := 3;
    StepTable[StepTc03Setup].StimulusId := 1;
    StepTable[StepTc03Setup].CheckIdx[1] := 1;
    StepTable[StepTc03Setup].TimeoutPT := T#12s;
    StepTable[StepTc03Setup].NextOnPass := StepTc03Trigger;
    StepTable[StepTc03Setup].NextOnFail := StepTc03Teardown;
    StepTable[StepTc03Setup].FailAction := E_TestFailAction.FAIL_CONTINUE;

    StepTable[StepTc03Trigger].Name := 'TCT3 Frequence fantome';
    StepTable[StepTc03Trigger].CaseId := 3;
    StepTable[StepTc03Trigger].StimulusId := 4;
    StepTable[StepTc03Trigger].CheckIdx[1] := 7;
    StepTable[StepTc03Trigger].CheckIdx[2] := 3;
    StepTable[StepTc03Trigger].CheckIdx[3] := 8;
    StepTable[StepTc03Trigger].TimeoutPT := T#4s;
    StepTable[StepTc03Trigger].NextOnPass := StepTc03Teardown;
    StepTable[StepTc03Trigger].NextOnFail := StepTc03Teardown;
    StepTable[StepTc03Trigger].FailAction := E_TestFailAction.FAIL_CONTINUE;

    StepTable[StepTc03Teardown].Name := 'TCT3 Teardown';
    StepTable[StepTc03Teardown].CaseId := 3;
    StepTable[StepTc03Teardown].StimulusId := 1;
    StepTable[StepTc03Teardown].CheckIdx[1] := 1;
    StepTable[StepTc03Teardown].TimeoutPT := T#12s;
    StepTable[StepTc03Teardown].NextOnPass := StepTc04Setup;
    StepTable[StepTc03Teardown].NextOnFail := StepTc04Setup;
    StepTable[StepTc03Teardown].FailAction := E_TestFailAction.FAIL_CONTINUE;

    // --- TC-T4 ---
    StepTable[StepTc04Setup].Name := 'TCT4 Setup saine';
    StepTable[StepTc04Setup].CaseId := 4;
    StepTable[StepTc04Setup].StimulusId := 1;
    StepTable[StepTc04Setup].CheckIdx[1] := 1;
    StepTable[StepTc04Setup].TimeoutPT := T#12s;
    StepTable[StepTc04Setup].NextOnPass := StepTc04Word1Tremie;
    StepTable[StepTc04Setup].NextOnFail := StepTc04Teardown;
    StepTable[StepTc04Setup].FailAction := E_TestFailAction.FAIL_CONTINUE;

    StepTable[StepTc04Word1Tremie].Name := 'TCT4 Mot 11111 Tremie';
    StepTable[StepTc04Word1Tremie].CaseId := 4;
    StepTable[StepTc04Word1Tremie].StimulusId := 5;
    StepTable[StepTc04Word1Tremie].CheckIdx[1] := 9;
    StepTable[StepTc04Word1Tremie].CheckIdx[2] := 10;
    StepTable[StepTc04Word1Tremie].CheckIdx[3] := 11;
    StepTable[StepTc04Word1Tremie].TimeoutPT := T#3s;
    StepTable[StepTc04Word1Tremie].NextOnPass := StepTc04Word2;
    StepTable[StepTc04Word1Tremie].NextOnFail := StepTc04Teardown;
    StepTable[StepTc04Word1Tremie].FailAction := E_TestFailAction.FAIL_CONTINUE;

    StepTable[StepTc04Word2].Name := 'TCT4 Mot 01111';
    StepTable[StepTc04Word2].CaseId := 4;
    StepTable[StepTc04Word2].StimulusId := 6;
    StepTable[StepTc04Word2].CheckIdx[1] := 9;
    StepTable[StepTc04Word2].TimeoutPT := T#3s;
    StepTable[StepTc04Word2].NextOnPass := StepTc04Word3;
    StepTable[StepTc04Word2].NextOnFail := StepTc04Teardown;
    StepTable[StepTc04Word2].FailAction := E_TestFailAction.FAIL_CONTINUE;

    StepTable[StepTc04Word3].Name := 'TCT4 Mot 00111';
    StepTable[StepTc04Word3].CaseId := 4;
    StepTable[StepTc04Word3].StimulusId := 7;
    StepTable[StepTc04Word3].CheckIdx[1] := 9;
    StepTable[StepTc04Word3].CheckIdx[2] := 14;
    StepTable[StepTc04Word3].CheckIdx[3] := 15;
    StepTable[StepTc04Word3].TimeoutPT := T#3s;
    StepTable[StepTc04Word3].NextOnPass := StepTc04Word4;
    StepTable[StepTc04Word3].NextOnFail := StepTc04Teardown;
    StepTable[StepTc04Word3].FailAction := E_TestFailAction.FAIL_CONTINUE;

    StepTable[StepTc04Word4].Name := 'TCT4 Mot 00011';
    StepTable[StepTc04Word4].CaseId := 4;
    StepTable[StepTc04Word4].StimulusId := 8;
    StepTable[StepTc04Word4].CheckIdx[1] := 9;
    StepTable[StepTc04Word4].TimeoutPT := T#3s;
    StepTable[StepTc04Word4].NextOnPass := StepTc04Word5;
    StepTable[StepTc04Word4].NextOnFail := StepTc04Teardown;
    StepTable[StepTc04Word4].FailAction := E_TestFailAction.FAIL_CONTINUE;

    StepTable[StepTc04Word5].Name := 'TCT4 Mot 00001';
    StepTable[StepTc04Word5].CaseId := 4;
    StepTable[StepTc04Word5].StimulusId := 9;
    StepTable[StepTc04Word5].CheckIdx[1] := 9;
    StepTable[StepTc04Word5].TimeoutPT := T#3s;
    StepTable[StepTc04Word5].NextOnPass := StepTc04Word6Maintenance;
    StepTable[StepTc04Word5].NextOnFail := StepTc04Teardown;
    StepTable[StepTc04Word5].FailAction := E_TestFailAction.FAIL_CONTINUE;

    StepTable[StepTc04Word6Maintenance].Name := 'TCT4 Mot 00000 Maintenance';
    StepTable[StepTc04Word6Maintenance].CaseId := 4;
    StepTable[StepTc04Word6Maintenance].StimulusId := 10;
    StepTable[StepTc04Word6Maintenance].CheckIdx[1] := 9;
    StepTable[StepTc04Word6Maintenance].CheckIdx[2] := 12;
    StepTable[StepTc04Word6Maintenance].CheckIdx[3] := 13;
    StepTable[StepTc04Word6Maintenance].TimeoutPT := T#3s;
    StepTable[StepTc04Word6Maintenance].NextOnPass := StepTc04Teardown;
    StepTable[StepTc04Word6Maintenance].NextOnFail := StepTc04Teardown;
    StepTable[StepTc04Word6Maintenance].FailAction := E_TestFailAction.FAIL_CONTINUE;

    StepTable[StepTc04Teardown].Name := 'TCT4 Teardown';
    StepTable[StepTc04Teardown].CaseId := 4;
    StepTable[StepTc04Teardown].StimulusId := 1;
    StepTable[StepTc04Teardown].CheckIdx[1] := 1;
    StepTable[StepTc04Teardown].TimeoutPT := T#12s;
    StepTable[StepTc04Teardown].NextOnPass := StepTc05Setup;
    StepTable[StepTc04Teardown].NextOnFail := StepTc05Setup;
    StepTable[StepTc04Teardown].FailAction := E_TestFailAction.FAIL_CONTINUE;

    // --- TC-T5 ---
    StepTable[StepTc05Setup].Name := 'TCT5 Setup saine';
    StepTable[StepTc05Setup].CaseId := 5;
    StepTable[StepTc05Setup].StimulusId := 1;
    StepTable[StepTc05Setup].CheckIdx[1] := 1;
    StepTable[StepTc05Setup].TimeoutPT := T#12s;
    StepTable[StepTc05Setup].NextOnPass := StepTc05Trigger;
    StepTable[StepTc05Setup].NextOnFail := StepTc05Teardown;
    StepTable[StepTc05Setup].FailAction := E_TestFailAction.FAIL_CONTINUE;

    StepTable[StepTc05Trigger].Name := 'TCT5 Mot incoherent force';
    StepTable[StepTc05Trigger].CaseId := 5;
    StepTable[StepTc05Trigger].StimulusId := 11;
    StepTable[StepTc05Trigger].CheckIdx[1] := 3;
    StepTable[StepTc05Trigger].CheckIdx[2] := 16;
    StepTable[StepTc05Trigger].CheckIdx[3] := 17;
    StepTable[StepTc05Trigger].CheckIdx[4] := 18;
    StepTable[StepTc05Trigger].TimeoutPT := T#5s;
    StepTable[StepTc05Trigger].NextOnPass := StepTc05Teardown;
    StepTable[StepTc05Trigger].NextOnFail := StepTc05Teardown;
    StepTable[StepTc05Trigger].FailAction := E_TestFailAction.FAIL_CONTINUE;

    StepTable[StepTc05Teardown].Name := 'TCT5 Teardown';
    StepTable[StepTc05Teardown].CaseId := 5;
    StepTable[StepTc05Teardown].StimulusId := 1;
    StepTable[StepTc05Teardown].CheckIdx[1] := 1;
    StepTable[StepTc05Teardown].TimeoutPT := T#12s;
    StepTable[StepTc05Teardown].NextOnPass := StepTc06Setup;
    StepTable[StepTc05Teardown].NextOnFail := StepTc06Setup;
    StepTable[StepTc05Teardown].FailAction := E_TestFailAction.FAIL_CONTINUE;

    // --- TC-T6 (instance isolée FB_Translation, voir fichier suite) ---
    StepTable[StepTc06Setup].Name := 'TCT6 Setup saine';
    StepTable[StepTc06Setup].CaseId := 6;
    StepTable[StepTc06Setup].StimulusId := 1;
    StepTable[StepTc06Setup].CheckIdx[1] := 1;
    StepTable[StepTc06Setup].TimeoutPT := T#12s;
    StepTable[StepTc06Setup].NextOnPass := StepTc06FullSpeed;
    StepTable[StepTc06Setup].NextOnFail := StepTc06Teardown;
    StepTable[StepTc06Setup].FailAction := E_TestFailAction.FAIL_CONTINUE;

    StepTable[StepTc06FullSpeed].Name := 'TCT6 Pleine vitesse sans PV';
    StepTable[StepTc06FullSpeed].CaseId := 6;
    StepTable[StepTc06FullSpeed].StimulusId := 12;
    StepTable[StepTc06FullSpeed].CheckIdx[1] := 19;
    StepTable[StepTc06FullSpeed].TimeoutPT := T#8s;
    StepTable[StepTc06FullSpeed].NextOnPass := StepTc06Slowdown;
    StepTable[StepTc06FullSpeed].NextOnFail := StepTc06Teardown;
    StepTable[StepTc06FullSpeed].FailAction := E_TestFailAction.FAIL_CONTINUE;

    StepTable[StepTc06Slowdown].Name := 'TCT6 Ralenti PV actif';
    StepTable[StepTc06Slowdown].CaseId := 6;
    StepTable[StepTc06Slowdown].StimulusId := 13;
    StepTable[StepTc06Slowdown].CheckIdx[1] := 20;
    StepTable[StepTc06Slowdown].TimeoutPT := T#8s;
    StepTable[StepTc06Slowdown].NextOnPass := StepTc06Teardown;
    StepTable[StepTc06Slowdown].NextOnFail := StepTc06Teardown;
    StepTable[StepTc06Slowdown].FailAction := E_TestFailAction.FAIL_CONTINUE;

    StepTable[StepTc06Teardown].Name := 'TCT6 Teardown';
    StepTable[StepTc06Teardown].CaseId := 6;
    StepTable[StepTc06Teardown].StimulusId := 1;
    StepTable[StepTc06Teardown].CheckIdx[1] := 1;
    StepTable[StepTc06Teardown].TimeoutPT := T#12s;
    StepTable[StepTc06Teardown].NextOnPass := 0;
    StepTable[StepTc06Teardown].NextOnFail := 0;
    StepTable[StepTc06Teardown].FailAction := E_TestFailAction.FAIL_CONTINUE;

    // 2. 🔒 VALIDATION — jouée UNE SEULE FOIS ici (les tables sont figées après
    //    construction, revalider chaque scan serait un coût inutile — 128 étapes max)
    ConfigError := FALSE;
ConfigErrorStepId := 0;
ConfigErrorCheckIdx := 0;
ConfigErrorMessage := '';

FOR Idx := 1 TO GVL_PLC_Tests_Const.MaxSteps DO
    IF StepTable[Idx].CaseId > 0 AND NOT ConfigError THEN
        IF StepTable[Idx].NextOnPass < 0 OR StepTable[Idx].NextOnPass > GVL_PLC_Tests_Const.MaxSteps THEN
            ConfigError := TRUE;
            ConfigErrorStepId := Idx;
            ConfigErrorMessage := 'NextOnPass hors limites';
        ELSIF StepTable[Idx].NextOnFail < 0 OR StepTable[Idx].NextOnFail > GVL_PLC_Tests_Const.MaxSteps THEN
            ConfigError := TRUE;
            ConfigErrorStepId := Idx;
            ConfigErrorMessage := 'NextOnFail hors limites';
        ELSIF StepTable[Idx].TimeoutPT <= T#0s THEN
            ConfigError := TRUE;
            ConfigErrorStepId := Idx;
            ConfigErrorMessage := 'TimeoutPT requis (> 0s)';
        ELSE
            FOR Jdx := 1 TO GVL_PLC_Tests_Const.MaxChecksPerStep DO
                Kdx := StepTable[Idx].CheckIdx[Jdx];
                IF Kdx > 0 AND NOT ConfigError THEN
                    IF Kdx > GVL_PLC_Tests_Const.MaxChecks THEN
                        ConfigError := TRUE;
                        ConfigErrorStepId := Idx;
                        ConfigErrorCheckIdx := Kdx;
                        ConfigErrorMessage := 'CheckIdx hors limites';
                    ELSE
                        // 📌 Périmètre restreint : seuls ces 3 Kind / 2 Mode sont supportés
                        CASE CheckTable[Kdx].Kind OF
                            E_TestCheckKind.BOOL_EQUAL:
                                IF CheckTable[Kdx].ProbeIdx < 1 OR CheckTable[Kdx].ProbeIdx > GVL_PLC_Tests_Const.MaxProbeBool THEN
                                    ConfigError := TRUE;
                                    ConfigErrorStepId := Idx;
                                    ConfigErrorCheckIdx := Kdx;
                                    ConfigErrorMessage := 'ProbeIdx BOOL hors limites';
                                END_IF;
                            E_TestCheckKind.WORD_MASK_NONE:
                                IF CheckTable[Kdx].ProbeIdx < 1 OR CheckTable[Kdx].ProbeIdx > GVL_PLC_Tests_Const.MaxProbeDint THEN
                                    ConfigError := TRUE;
                                    ConfigErrorStepId := Idx;
                                    ConfigErrorCheckIdx := Kdx;
                                    ConfigErrorMessage := 'ProbeIdx DINT hors limites';
                                END_IF;
                            E_TestCheckKind.REAL_IN_RANGE:
                                IF CheckTable[Kdx].ProbeIdx < 1 OR CheckTable[Kdx].ProbeIdx > GVL_PLC_Tests_Const.MaxProbeReal THEN
                                    ConfigError := TRUE;
                                    ConfigErrorStepId := Idx;
                                    ConfigErrorCheckIdx := Kdx;
                                    ConfigErrorMessage := 'ProbeIdx REAL hors limites';
                                END_IF;
                        ELSE
                            ConfigError := TRUE;
                            ConfigErrorStepId := Idx;
                            ConfigErrorCheckIdx := Kdx;
                            ConfigErrorMessage := 'Kind non supporte par ce moteur dedie';
                        END_CASE;

                        IF NOT ConfigError THEN
                            IF CheckTable[Kdx].Mode <> E_TestCheckMode.CHECK_WAIT_UNTIL AND CheckTable[Kdx].Mode <> E_TestCheckMode.CHECK_INSTANT THEN
                                ConfigError := TRUE;
                                ConfigErrorStepId := Idx;
                                ConfigErrorCheckIdx := Kdx;
                                ConfigErrorMessage := 'Mode non supporte par ce moteur dedie';
                            END_IF;
                        END_IF;
                    END_IF;
                END_IF;
            END_FOR;
        END_IF;
    END_IF;
END_FOR;

// Cohérence CaseTable[1..6] <-> StepTable (chaque case doit démarrer sur SON setup)
IF NOT ConfigError THEN
    FOR Idx := 1 TO 6 DO
        IF CaseTable[Idx].FirstStep < 1 OR CaseTable[Idx].FirstStep > GVL_PLC_Tests_Const.MaxSteps THEN
            ConfigError := TRUE;
            ConfigErrorStepId := CaseTable[Idx].FirstStep;
            ConfigErrorMessage := 'CaseTable.FirstStep hors limites';
        ELSIF StepTable[CaseTable[Idx].FirstStep].CaseId <> Idx THEN
            ConfigError := TRUE;
            ConfigErrorStepId := CaseTable[Idx].FirstStep;
            ConfigErrorMessage := 'CaseTable.FirstStep ne pointe pas vers SON case';
        END_IF;
    END_FOR;
END_IF;

// 🔒 Validation structurelle complémentaire : stimulus connu, étape utile,
// cibles configurées et changement de case réservé au teardown (Pass=Fail).
IF NOT ConfigError THEN
    FOR Idx := 1 TO GVL_PLC_Tests_Const.MaxSteps DO
        IF StepTable[Idx].CaseId > 0 AND NOT ConfigError THEN
            IF StepTable[Idx].StimulusId < 0 OR StepTable[Idx].StimulusId > 13 THEN
                ConfigError := TRUE; ConfigErrorStepId := Idx;
                ConfigErrorMessage := 'StimulusId hors plage Translation 0..13';
            END_IF;
            HasCheck := FALSE;
            FOR Jdx := 1 TO GVL_PLC_Tests_Const.MaxChecksPerStep DO
                HasCheck := HasCheck OR (StepTable[Idx].CheckIdx[Jdx] > 0);
            END_FOR;
            IF NOT HasCheck AND StepTable[Idx].DwellPT <= T#0s THEN
                ConfigError := TRUE; ConfigErrorStepId := Idx;
                ConfigErrorMessage := 'Etape sans check ni dwell explicite';
            END_IF;
            // 🔒 Branches imbriquées : aucun StepTable[0], sans supposer AND court-circuité.
            IF StepTable[Idx].NextOnPass > 0 THEN
                Kdx := StepTable[Idx].NextOnPass;
                IF StepTable[Kdx].CaseId = 0 THEN
                    ConfigError := TRUE; ConfigErrorStepId := Idx;
                    ConfigErrorMessage := 'NextOnPass vise une etape non configuree';
                END_IF;
            END_IF;
            IF StepTable[Idx].NextOnFail > 0 AND NOT ConfigError THEN
                Kdx := StepTable[Idx].NextOnFail;
                IF StepTable[Kdx].CaseId = 0 THEN
                    ConfigError := TRUE; ConfigErrorStepId := Idx;
                    ConfigErrorMessage := 'NextOnFail vise une etape non configuree';
                ELSIF StepTable[Kdx].CaseId <> StepTable[Idx].CaseId THEN
                    IF StepTable[Idx].NextOnPass <> StepTable[Idx].NextOnFail THEN
                        ConfigError := TRUE; ConfigErrorStepId := Idx;
                        ConfigErrorMessage := 'Echec quitte le case sans teardown commun';
                    END_IF;
                END_IF;
            END_IF;
        END_IF;
    END_FOR;
END_IF;

// 🔁 Chaque chemin nominal Case→fin doit sortir en <= MaxSteps transitions.
IF NOT ConfigError THEN
    FOR Idx := 1 TO 6 DO
        WalkStep := CaseTable[Idx].FirstStep;
        FOR WalkIdx := 1 TO GVL_PLC_Tests_Const.MaxSteps DO
            IF WalkStep = 0 THEN EXIT; END_IF;
            // 🔒 Valider la borne avant de déréférencer WalkStep.
            IF WalkStep < 1 OR WalkStep > GVL_PLC_Tests_Const.MaxSteps THEN
                ConfigError := TRUE; ConfigErrorStepId := WalkStep;
                ConfigErrorMessage := 'Chemin nominal hors limites';
                EXIT;
            END_IF;
            IF StepTable[WalkStep].CaseId = 0 THEN
                ConfigError := TRUE; ConfigErrorStepId := WalkStep;
                ConfigErrorMessage := 'Chemin nominal non configure';
                EXIT;
            END_IF;
            WalkStep := StepTable[WalkStep].NextOnPass;
        END_FOR;
        IF WalkStep <> 0 AND NOT ConfigError THEN
            ConfigError := TRUE; ConfigErrorStepId := WalkStep;
            ConfigErrorMessage := 'Cycle nominal ou chemin sans sortie';
        END_IF;
    END_FOR;
END_IF;

    Ready := NOT ConfigError;
    Built := TRUE;
END_IF;

(* ---- FB_TranslationTestRuntime.st ---- *)
// ═══════════════════════════════════════════════════════════════
// 🧪 FB_TranslationTestRuntime — Cycle de vie protégé Translation M3
// ───────────────────────────────────────────────────────────────
// 🎯 Responsabilité UNIQUE : posséder le lifecycle atomique du run :
//    IDLE → RUN → CLEANUP → WAIT_NEUTRAL → VERIFY → TERMINAL.
// 🔒 Aucun terminal n'est publié avant neutralité confirmée.
// ═══════════════════════════════════════════════════════════════

FUNCTION_BLOCK PUBLIC FB_TranslationTestRuntime
VAR_INPUT
    Start   : BOOL;
    Abort   : BOOL;
    CaseId  : INT;
    PlanConfigError         : BOOL;
    PlanConfigErrorStepId   : INT;
    PlanConfigErrorCheckIdx : INT;
    PlanConfigErrorMessage  : STRING(160);
    SimulationModeActive    : BOOL;
    SimGateOk               : BOOL;
    NeutralConfirmed        : BOOL; // Neutralité réellement appliquée au scan précédent
    WatchdogLimitMs         : DINT := 180000; // Paramétrable pour autotest du framework
    CleanupTimeoutScans     : INT := 20;      // Délai max de confirmation du neutre
END_VAR
VAR_IN_OUT
    StepTable  : ARRAY[1..GVL_PLC_Tests_Const.MaxSteps]      OF ST_TestStepConfig;
    CheckTable : ARRAY[1..GVL_PLC_Tests_Const.MaxChecks]     OF ST_TestCheckConfig;
    CaseTable  : ARRAY[1..GVL_PLC_Tests_Const.MaxTestCases]  OF ST_TestCaseConfig;
    ProbeBool  : ARRAY[1..GVL_PLC_Tests_Const.MaxProbeBool]  OF BOOL;
    ProbeDint  : ARRAY[1..GVL_PLC_Tests_Const.MaxProbeDint]  OF DINT;
    ProbeReal  : ARRAY[1..GVL_PLC_Tests_Const.MaxProbeReal]  OF REAL;
    Report     : ST_TestSuiteReport;
    Result     : ST_TranslationTestResult;
END_VAR
VAR_OUTPUT
    Busy                : BOOL;
    Done                : BOOL;
    AnyFailed           : BOOL;
    ActiveStimulusId    : INT;
    StepElapsed         : TIME;
    TerminalState       : E_TestTerminalState;
    ConfigError         : BOOL;
    ConfigErrorStepId   : INT;
    ConfigErrorCheckIdx : INT;
    ErrorCode           : INT;
    ErrorMessage        : STRING(160);
    StartRejected       : BOOL; // Impulsion : Start reçu hors IDLE/TERMINAL
    CleanupRequest      : BOOL; // Niveau : imposer le vecteur neutre complet
END_VAR
VAR CONSTANT
    RuntimeIdle        : INT := 0;
    RuntimeRun         : INT := 10;
    RuntimeCleanup     : INT := 20;
    RuntimeWaitNeutral : INT := 30;
    RuntimeVerify      : INT := 40;
    RuntimeTerminal    : INT := 50;
END_VAR
VAR
    instFixture   : FB_TranslationTestFixture;
    instExecutor  : FB_TranslationStepExecutor;
    instFinalizer : FB_TranslationReportFinalizer;
    StartTrig     : R_TRIG;
    RuntimeState  : INT := 0;
    ExecutorStart : BOOL;
    ExecutorAbort : BOOL;
    RunStartPulse : BOOL;
    FinalizePulse : BOOL;
    PendingTerminalState : E_TestTerminalState;
    PendingErrorCode     : INT;
    PendingErrorMessage  : STRING(160);
    SuiteElapsed         : TIME;
    NeutralWaitScans     : INT;
    CleanupElapsedScans  : INT;
END_VAR
// === IMPLEMENTATION ===
StartTrig(CLK := Start);
StartRejected := FALSE;
ExecutorStart := FALSE;
ExecutorAbort := FALSE;
RunStartPulse := FALSE;
FinalizePulse := FALSE;
CleanupRequest := (RuntimeState = RuntimeCleanup)
               OR (RuntimeState = RuntimeWaitNeutral)
               OR (RuntimeState = RuntimeVerify);

// 🎮 Un Start pendant un run/cleanup est refusé sans modifier le run actif.
IF StartTrig.Q AND RuntimeState <> RuntimeIdle AND RuntimeState <> RuntimeTerminal THEN
    StartRejected := TRUE;
END_IF;

// 🚪 Fixture appelée CHAQUE scan : son R_TRIG interne est ainsi toujours réarmé.
instFixture(CheckRequested := StartTrig.Q,
            SimulationModeActive := SimulationModeActive,
            SimGateOk := SimGateOk);

// 🟢 Nouveau run accepté depuis IDLE ou TERMINAL.
IF StartTrig.Q AND (RuntimeState = RuntimeIdle OR RuntimeState = RuntimeTerminal) THEN
    RunStartPulse := TRUE;
    Done := FALSE;
    SuiteElapsed := T#0s;
    NeutralWaitScans := 0;
    CleanupElapsedScans := 0;
    PendingTerminalState := E_TestTerminalState.TEST_TERMINAL_NONE;
    PendingErrorCode := 0;
    PendingErrorMessage := '';

    IF PlanConfigError THEN
        PendingTerminalState := E_TestTerminalState.TEST_TERMINAL_CONFIG_ERROR;
        PendingErrorCode := 1002;
        PendingErrorMessage := CONCAT('Table invalide : ', PlanConfigErrorMessage);
        RuntimeState := RuntimeCleanup;
    ELSIF CaseId < 0 OR CaseId > 6 THEN
        PendingTerminalState := E_TestTerminalState.TEST_TERMINAL_CONFIG_ERROR;
        PendingErrorCode := 1001;
        PendingErrorMessage := 'CaseId invalide (attendu 0..6)';
        RuntimeState := RuntimeCleanup;
    ELSIF instFixture.FixtureFailed THEN
        PendingTerminalState := E_TestTerminalState.TEST_TERMINAL_PRECONDITION_FAILED;
        PendingErrorCode := 1010;
        PendingErrorMessage := CONCAT('PRECONDITION_FAILED : ', instFixture.FailReason);
        RuntimeState := RuntimeCleanup;
    ELSE
        ExecutorStart := TRUE;
        RuntimeState := RuntimeRun;
    END_IF;
END_IF;

// 🛡️ Causes de sortie du RUN : watchdog > gate perdue > abort opérateur.
IF RuntimeState = RuntimeRun THEN
    SuiteElapsed := SuiteElapsed + UDINT_TO_TIME(INT_TO_UDINT(GVL_PLC_Tests_Const.TaskCycleMs));
    IF SuiteElapsed >= DINT_TO_TIME(WatchdogLimitMs) THEN
        ExecutorAbort := TRUE;
        PendingTerminalState := E_TestTerminalState.TEST_TERMINAL_WATCHDOG_TIMEOUT;
        PendingErrorCode := 1020;
        PendingErrorMessage := 'Watchdog suite Translation expire';
    ELSIF NOT SimulationModeActive OR NOT SimGateOk THEN
        ExecutorAbort := TRUE;
        PendingTerminalState := E_TestTerminalState.TEST_TERMINAL_PRECONDITION_FAILED;
        PendingErrorCode := 1011;
        PendingErrorMessage := 'Gate Translation perdue pendant le run';
    ELSIF Abort THEN
        ExecutorAbort := TRUE;
        PendingTerminalState := E_TestTerminalState.TEST_TERMINAL_ABORTED;
        PendingErrorCode := 1030;
        PendingErrorMessage := 'Abandon operateur';
    END_IF;
END_IF;

// 🪜 L'exécuteur ne possède que les étapes, jamais le terminal public.
instExecutor(
    Start := ExecutorStart,
    Abort := ExecutorAbort,
    CaseId := CaseId,
    StepTable := StepTable,
    CheckTable := CheckTable,
    CaseTable := CaseTable,
    ProbeBool := ProbeBool,
    ProbeDint := ProbeDint,
    ProbeReal := ProbeReal
);

IF RuntimeState = RuntimeRun AND instExecutor.RunDone THEN
    IF PendingTerminalState = E_TestTerminalState.TEST_TERMINAL_NONE THEN
        PendingTerminalState := instExecutor.TerminalState;
        IF instExecutor.ConfigError THEN
            PendingErrorCode := 1003;
            PendingErrorMessage := 'Garde-fou runtime : transition invalide';
        END_IF;
    END_IF;
    RuntimeState := RuntimeCleanup;
    NeutralWaitScans := 0;
END_IF;

// 🧹 Tous les chemins imposent au moins deux scans complets au neutre.
IF RuntimeState = RuntimeCleanup THEN
    CleanupRequest := TRUE;
    NeutralWaitScans := 0;
    CleanupElapsedScans := 0;
    RuntimeState := RuntimeWaitNeutral;
ELSIF RuntimeState = RuntimeWaitNeutral THEN
    CleanupRequest := TRUE;
    NeutralWaitScans := NeutralWaitScans + 1;
    CleanupElapsedScans := CleanupElapsedScans + 1;
    IF NeutralWaitScans >= 2 THEN
        RuntimeState := RuntimeVerify;
    END_IF;
ELSIF RuntimeState = RuntimeVerify THEN
    CleanupRequest := TRUE;
    CleanupElapsedScans := CleanupElapsedScans + 1;
    IF NeutralConfirmed THEN
        FinalizePulse := TRUE;
        RuntimeState := RuntimeTerminal;
        Done := TRUE;
    ELSIF CleanupElapsedScans >= CleanupTimeoutScans THEN
        PendingTerminalState := E_TestTerminalState.TEST_TERMINAL_CONFIG_ERROR;
        PendingErrorCode := 1040;
        PendingErrorMessage := 'Cleanup Translation non confirme';
        FinalizePulse := TRUE;
        RuntimeState := RuntimeTerminal;
        Done := TRUE;
    END_IF;
END_IF;

// 📊 Le rapport consomme directement chaque verdict, même consécutif.
instFinalizer(
    RunStart := RunStartPulse,
    RequestedCaseId := CaseId,
    Busy := (RuntimeState = RuntimeRun),
    StepVerdict := instExecutor.StepVerdict,
    StepId := instExecutor.VerdictStepId,
    StepCaseId := instExecutor.VerdictCaseId,
    StepPassed := instExecutor.VerdictPassed,
    StepFailReason := instExecutor.VerdictFailReason,
    StepFailedCheckIdx := instExecutor.VerdictFailedCheckIdx,
    StepDuration := instExecutor.VerdictDuration,
    StepObservedBool := instExecutor.VerdictObservedBool,
    StepObservedDint := instExecutor.VerdictObservedDint,
    StepObservedReal := instExecutor.VerdictObservedReal,
    Finalize := FinalizePulse,
    TerminalState := PendingTerminalState,
    ErrorCode := PendingErrorCode,
    ErrorMessage := PendingErrorMessage,
    StepTable := StepTable,
    CaseTable := CaseTable,
    Report := Report,
    Result := Result
);

// 📤 Publication : Busy inclut cleanup ; aucun stimulus métier hors RUN.
Busy := (RuntimeState = RuntimeRun)
     OR (RuntimeState = RuntimeCleanup)
     OR (RuntimeState = RuntimeWaitNeutral)
     OR (RuntimeState = RuntimeVerify);
IF RuntimeState = RuntimeRun THEN
    ActiveStimulusId := instExecutor.ActiveStimulusId;
ELSE
    ActiveStimulusId := 0;
END_IF;
StepElapsed := instExecutor.StepElapsed;
TerminalState := Result.TerminalState;
AnyFailed := Result.AnyFailed;
ConfigError := PlanConfigError OR instExecutor.ConfigError;
IF PlanConfigError THEN
    ConfigErrorStepId := PlanConfigErrorStepId;
    ConfigErrorCheckIdx := PlanConfigErrorCheckIdx;
ELSE
    ConfigErrorStepId := instExecutor.ConfigErrorStepId;
    ConfigErrorCheckIdx := 0;
END_IF;
ErrorCode := Result.ErrorCode;
ErrorMessage := Result.ErrorMessage;
